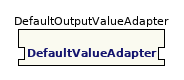
      [picture p48: application _05_Adapter.Ex4b]
      FBS
        DefaultOutputValueAdapter : DefaultValueAdapter;
      END_FBS
    END_SUBAPPLICATION
  END_APPLICATION
  DEVICE RaspberryPI : (MGR_ID := "localhost:61499")
    {SET_ATTRIBUTE(Profile, HOLOBLOC)}
    RESOURCE EMB_RES : 
    END_RESOURCE
  END_DEVICE
END_SYSTEM
